FUNCTION_BLOCK ASSEMBLE_AQ_FROM_AX (* this Function combines the 2 AX (BOOL) adapters to a AQ (QUARTER) *)
  (* Standard: 61499-2; Description: Copyright (c) 2026 HR Agrartechnik GmbH This program and the accompanying materials are made available under the terms of the Eclipse Public License 2.0 which is available at https://www.eclipse.org/legal/epl-2.0/ SPDX-License-Identifier: EPL-2.0 *)
  (* Version 1.0, 2026-11-13, Franz Höpfinger, HR Agrartechnik GmbH, Initial Version - Luecke in der Adapter-Familie geschlossen *)
  PACKAGE adapter::assembling;
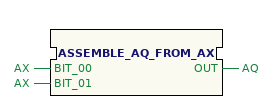
  SOCKETS
    BIT_00 : adapter::types::unidirectional::AX; (* Bool Bit 0 *)
    BIT_01 : adapter::types::unidirectional::AX; (* Bool Bit 1 *)
  END_SOCKETS
  PLUGS
    OUT : adapter::types::unidirectional::AQ; (* QUARTER Output (Bit 0 und 1) *)
  END_PLUGS
END_FUNCTION_BLOCK
